(* IEC 61131-3 sources: kns-pump-station/tests/GVLs, 3 files *)

(* ---- GVL_TestsInfra.gvl.st ---- *)
// Назначение: экземпляры наборов тестов команды К3 (сгенерированный слой, полевой слой, журнал, сводка тревог).
//             Объявление регистрирует набор в coUnit; {attribute 'linkalways'} обязателен — без него
//             компилятор выбросит GVL, на которую никто не ссылается, и наборы молча пропадут.
// Автор:      kr0nsch
// Версия:     0.1.0
// Документ:   docs/DESIGN.md, раздел 14.1
{attribute 'qualified_only'}
{attribute 'linkalways'}
VAR_GLOBAL
    fbVfdAdapterCondTest : FB_VfdAdapter_Cond_Test;   // 8.2
    fbEventLogTest       : FB_EventLog_Test;          // 9.1
    fbEventLogCsvTest    : FB_EventLogCsv_Test;       // 9.2 (многоцикловые, CAA File)
    fbUtcToIsoTest       : FB_F_UtcToIso_Test;        // 9.2
    fbAlarmCodeTest      : FB_F_AlarmCode_Test;       // 9.2
    fbAlarmSummaryTest   : FB_AlarmSummary_Test;      // 9.3
    fbDeviceAuditTest    : FB_DeviceAudit_Test;       // 9.3
    fbPlcStartAdoptionTest : FB_PlcStartAdoption_Test;  // 4.6, 7: подхват насоса в порядке PRG_Devices
    fbFieldOwenTest : FB_FieldOwen_Test;      // 8.4: функции полевого слоя ОВЕН (сборка targets/plc210)
END_VAR

(* ---- GVL_TestsModel.gvl.st ---- *)
// Назначение: экземпляры наборов тестов модели, имитации и часов (команда К2). Набор coUnit
//             регистрируется объявлением экземпляра; {attribute 'linkalways'} обязателен — иначе
//             компилятор выбросит GVL, на которую никто не ссылается, и наборы молча пропадут
//             (решение F-01 plc-process-lib, docs/TESTING.md библиотеки).
// Автор:      kr0nsch
// Версия:     0.1.0
// Документ:   docs/DESIGN.md, разделы 11.3, 14.1
{attribute 'qualified_only'}
{attribute 'linkalways'}
VAR_GLOBAL
    fbScaledClockTest     : FB_ScaledClock_Test;
    fbInflowProfileTest   : FB_InflowProfile_Test;
    fbStormGeneratorTest  : FB_StormGenerator_Test;
    fbTankModelTest       : FB_TankModel_Test;
    fbHydraulicSolverTest : FB_HydraulicSolver_Test;
    fbVfdSimTest          : FB_VfdSim_Test;
    fbPlantModelTest      : FB_PlantModel_Test;
END_VAR

(* ---- GVL_TestsStation.gvl.st ---- *)
// Назначение: экземпляры наборов тестов логики станции (команда «логика станции», DESIGN 14.1).
//             Объявление регистрирует набор в coUnit; {attribute 'linkalways'} обязателен — без него
//             компилятор выбросит GVL, на которую никто не ссылается, и наборы молча пропадут.
// Автор:      kr0nsch
// Версия:     0.1.0
// Документ:   docs/DESIGN.md, раздел 14.1
{attribute 'qualified_only'}
{attribute 'linkalways'}
VAR_GLOBAL
    fbStationModeTest          : FB_StationMode_Test;           // 6.1
    fbControlSelectorTest      : FB_ControlSelector_Test;       // 6.2
    fbLevelControlSteppedTest  : FB_LevelControlStepped_Test;   // 6.3
    fbLevelControlPidTest      : FB_LevelControlPid_Test;       // 6.4
    fbPumpRotationTest         : FB_PumpRotation_Test;          // 6.5
    fbAtsTest                  : FB_Ats_Test;                   // 6.6
    fbProtectionsTest          : FB_Protections_Test;           // 6.7
    fbPumpProtectionTest       : FB_PumpProtection_Test;        // 6.8
    fbPowerRestoreTest         : FB_PowerRestore_Test;          // 6.9
    fbVentilationTest          : FB_Ventilation_Test;           // 6.10
    fbStationAlarmsTest        : FB_StationAlarms_Test;         // 6.11
    fbAnnunciatorTest          : FB_Annunciator_Test;           // 6.12
    fbStationCfgCheckTest      : FB_F_StationCfgCheck_Test;     // 6.13
    fbStationCoreTest          : FB_StationCore_Test;           // 6.15, раздел 7
END_VAR
